// Mitsubishi GX Works2 project: v2(working)   PLC: FX3U/FX3UC

PROGRAM MAIN
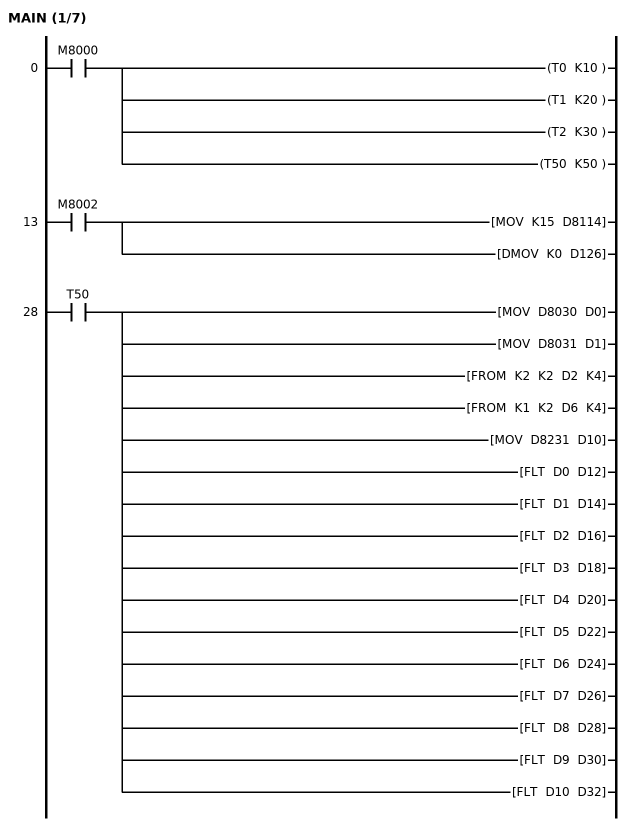
0     LD      M8000
      OUT     T0 K10
      OUT     T1 K20
      OUT     T2 K30
      OUT     T50 K50
13    LD      M8002
      MOV     K15 D8114
      DMOV    K0 D126
28    LD      T50
      MOV     D8030 D0
      MOV     D8031 D1
      FROM    K2 K2 D2 K4
      FROM    K1 K2 D6 K4
      MOV     D8231 D10
      FLT     D0 D12
      FLT     D1 D14
      FLT     D2 D16
      FLT     D3 D18
      FLT     D4 D20
      FLT     D5 D22
      FLT     D6 D24
      FLT     D7 D26
      FLT     D8 D28
      FLT     D9 D30
      FLT     D10 D32
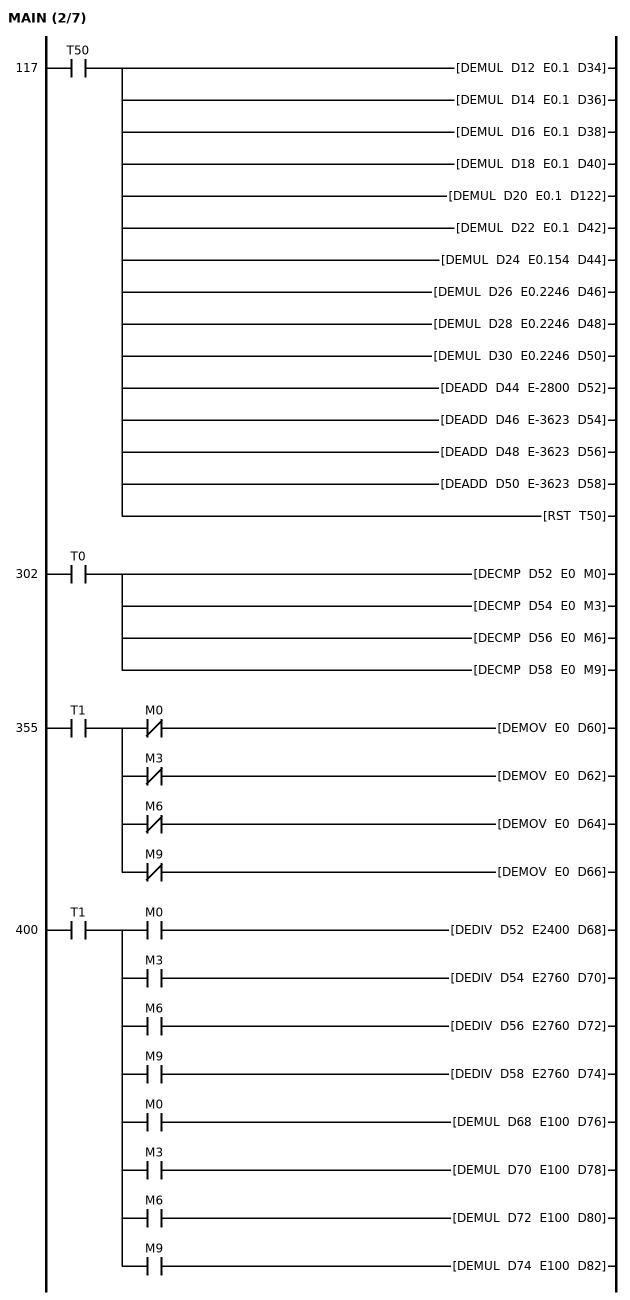
117   LD      T50
      DEMUL   D12 E0.1 D34
      DEMUL   D14 E0.1 D36
      DEMUL   D16 E0.1 D38
      DEMUL   D18 E0.1 D40
      DEMUL   D20 E0.1 D122
      DEMUL   D22 E0.1 D42
      DEMUL   D24 E0.154 D44
      DEMUL   D26 E0.2246 D46
      DEMUL   D28 E0.2246 D48
      DEMUL   D30 E0.2246 D50
      DEADD   D44 E-2800 D52
      DEADD   D46 E-3623 D54
      DEADD   D48 E-3623 D56
      DEADD   D50 E-3623 D58
      RST     T50
302   LD      T0
      DECMP   D52 E0 M0
      DECMP   D54 E0 M3
      DECMP   D56 E0 M6
      DECMP   D58 E0 M9
355   LD      T1
      MPS
      ANI     M0
      DEMOV   E0 D60
      MRD
      ANI     M3
      DEMOV   E0 D62
      MRD
      ANI     M6
      DEMOV   E0 D64
      MPP
      ANI     M9
      DEMOV   E0 D66
400   LD      T1
      MPS
      AND     M0
      DEDIV   D52 E2400 D68
      MRD
      AND     M3
      DEDIV   D54 E2760 D70
      MRD
      AND     M6
      DEDIV   D56 E2760 D72
      MRD
      AND     M9
      DEDIV   D58 E2760 D74
      MRD
      AND     M0
      DEMUL   D68 E100 D76
      MRD
      AND     M3
      DEMUL   D70 E100 D78
      MRD
      AND     M6
      DEMUL   D72 E100 D80
      MPP
      AND     M9
      DEMUL   D74 E100 D82
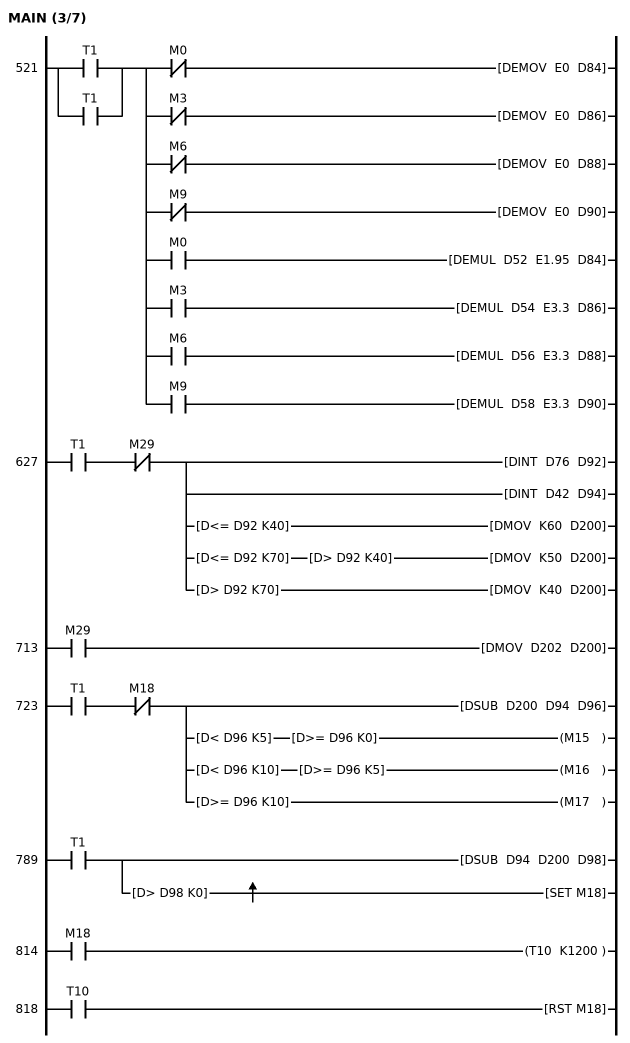
521   LD      T1
      OR      T1
      MPS
      ANI     M0
      DEMOV   E0 D84
      MRD
      ANI     M3
      DEMOV   E0 D86
      MRD
      ANI     M6
      DEMOV   E0 D88
      MRD
      ANI     M9
      DEMOV   E0 D90
      MRD
      AND     M0
      DEMUL   D52 E1.95 D84
      MRD
      AND     M3
      DEMUL   D54 E3.3 D86
      MRD
      AND     M6
      DEMUL   D56 E3.3 D88
      MPP
      AND     M9
      DEMUL   D58 E3.3 D90
627   LD      T1
      ANI     M29
      DINT    D76 D92
      DINT    D42 D94
      MPS
      ANDD<=  D92 K40
      DMOV    K60 D200
      MRD
      ANDD<=  D92 K70
      ANDD>   D92 K40
      DMOV    K50 D200
      MPP
      ANDD>   D92 K70
      DMOV    K40 D200
713   LD      M29
      DMOV    D202 D200
723   LD      T1
      ANI     M18
      DSUB    D200 D94 D96
      MPS
      ANDD<   D96 K5
      ANDD>=  D96 K0
      OUT     M15
      MRD
      ANDD<   D96 K10
      ANDD>=  D96 K5
      OUT     M16
      MPP
      ANDD>=  D96 K10
      OUT     M17
789   LD      T1
      DSUB    D94 D200 D98
      ANDD>   D98 K0
      MEP
      SET     M18
814   LD      M18
      OUT     T10 K1200
818   LD      T10
      RST     M18
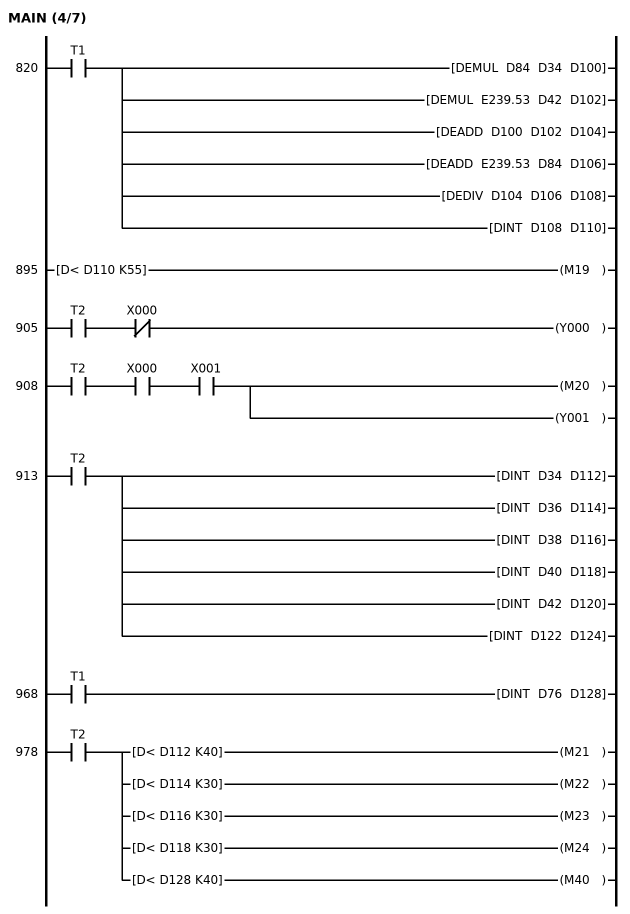
820   LD      T1
      DEMUL   D84 D34 D100
      DEMUL   E239.53 D42 D102
      DEADD   D100 D102 D104
      DEADD   E239.53 D84 D106
      DEDIV   D104 D106 D108
      DINT    D108 D110
895   LDD<    D110 K55
      OUT     M19
905   LD      T2
      ANI     X000
      OUT     Y000
908   LD      T2
      AND     X000
      AND     X001
      OUT     M20
      OUT     Y001
913   LD      T2
      DINT    D34 D112
      DINT    D36 D114
      DINT    D38 D116
      DINT    D40 D118
      DINT    D42 D120
      DINT    D122 D124
968   LD      T1
      DINT    D76 D128
978   LD      T2
      MPS
      ANDD<   D112 K40
      OUT     M21
      MRD
      ANDD<   D114 K30
      OUT     M22
      MRD
      ANDD<   D116 K30
      OUT     M23
      MRD
      ANDD<   D118 K30
      OUT     M24
      MPP
      ANDD<   D128 K40
      OUT     M40
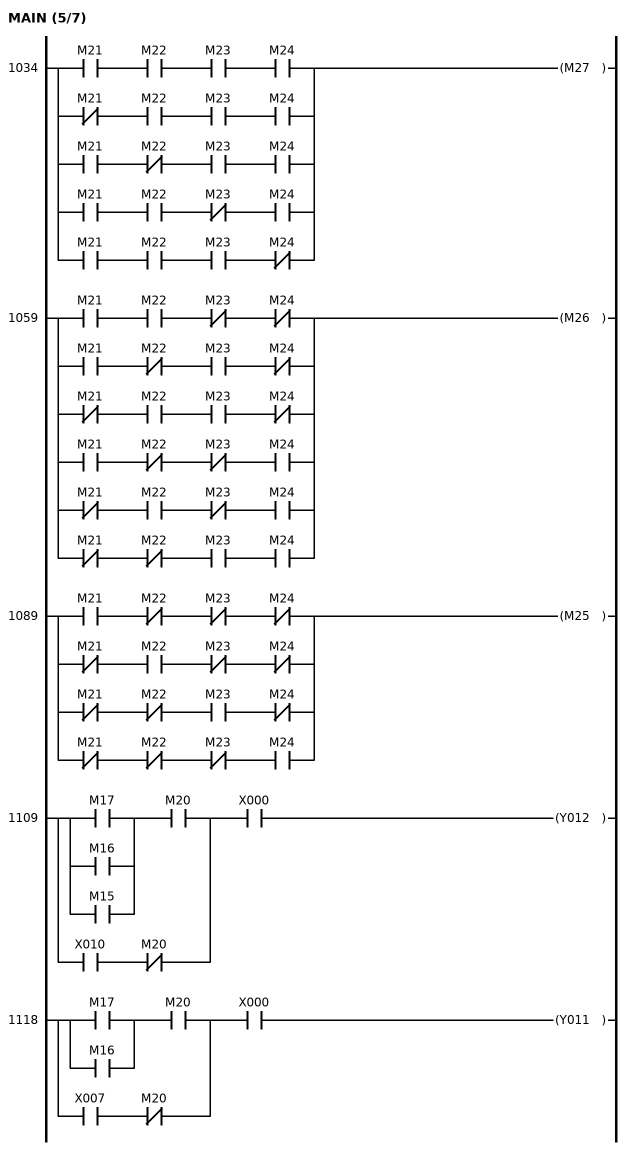
1034  LD      M21
      AND     M22
      AND     M23
      AND     M24
      LDI     M21
      AND     M22
      AND     M23
      AND     M24
      ORB
      LD      M21
      ANI     M22
      AND     M23
      AND     M24
      ORB
      LD      M21
      AND     M22
      ANI     M23
      AND     M24
      ORB
      LD      M21
      AND     M22
      AND     M23
      ANI     M24
      ORB
      OUT     M27
1059  LD      M21
      AND     M22
      ANI     M23
      ANI     M24
      LD      M21
      ANI     M22
      AND     M23
      ANI     M24
      ORB
      LDI     M21
      AND     M22
      AND     M23
      ANI     M24
      ORB
      LD      M21
      ANI     M22
      ANI     M23
      AND     M24
      ORB
      LDI     M21
      AND     M22
      ANI     M23
      AND     M24
      ORB
      LDI     M21
      ANI     M22
      AND     M23
      AND     M24
      ORB
      OUT     M26
1089  LD      M21
      ANI     M22
      ANI     M23
      ANI     M24
      LDI     M21
      AND     M22
      ANI     M23
      ANI     M24
      ORB
      LDI     M21
      ANI     M22
      AND     M23
      ANI     M24
      ORB
      LDI     M21
      ANI     M22
      ANI     M23
      AND     M24
      ORB
      OUT     M25
1109  LD      M17
      OR      M16
      OR      M15
      AND     M20
      LD      X010
      ANI     M20
      ORB
      AND     X000
      OUT     Y012
1118  LD      M17
      OR      M16
      AND     M20
      LD      X007
      ANI     M20
      ORB
      AND     X000
      OUT     Y011
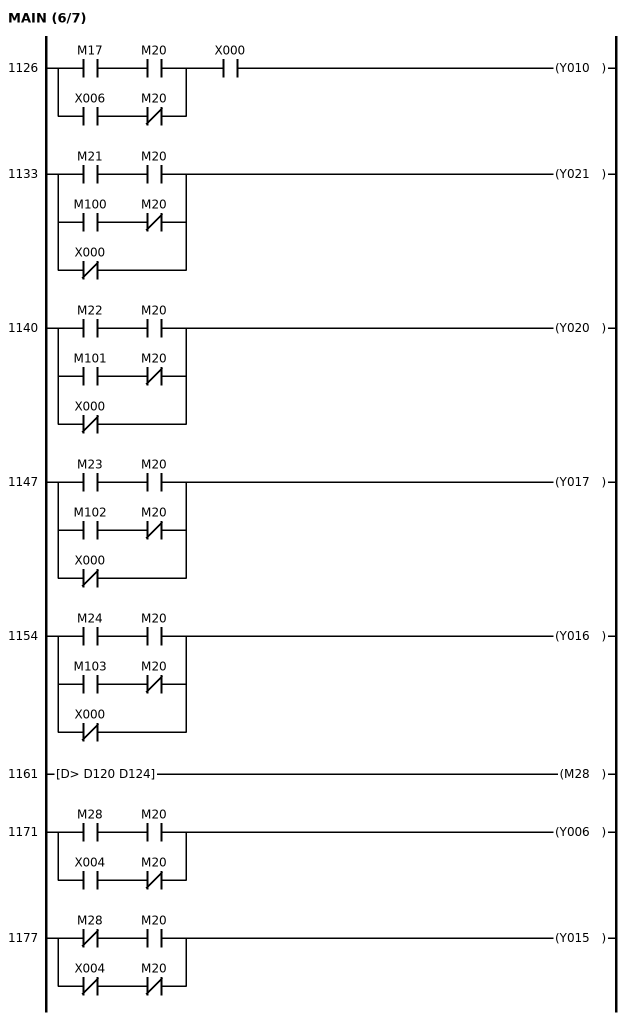
1126  LD      M17
      AND     M20
      LD      X006
      ANI     M20
      ORB
      AND     X000
      OUT     Y010
1133  LD      M21
      AND     M20
      LD      M100
      ANI     M20
      ORB
      ORI     X000
      OUT     Y021
1140  LD      M22
      AND     M20
      LD      M101
      ANI     M20
      ORB
      ORI     X000
      OUT     Y020
1147  LD      M23
      AND     M20
      LD      M102
      ANI     M20
      ORB
      ORI     X000
      OUT     Y017
1154  LD      M24
      AND     M20
      LD      M103
      ANI     M20
      ORB
      ORI     X000
      OUT     Y016
1161  LDD>    D120 D124
      OUT     M28
1171  LD      M28
      AND     M20
      LD      X004
      ANI     M20
      ORB
      OUT     Y006
1177  LDI     M28
      AND     M20
      LDI     X004
      ANI     M20
      ORB
      OUT     Y015
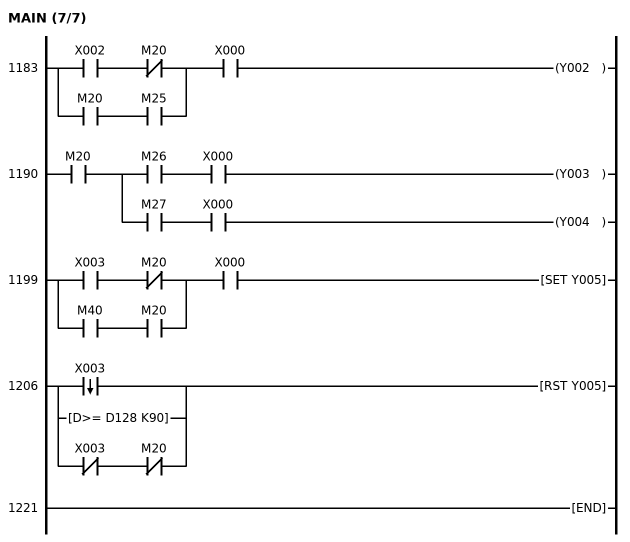
1183  LD      X002
      ANI     M20
      LD      M20
      AND     M25
      ORB
      AND     X000
      OUT     Y002
1190  LD      M20
      MPS
      AND     M26
      AND     X000
      OUT     Y003
      MPP
      AND     M27
      AND     X000
      OUT     Y004
1199  LD      X003
      ANI     M20
      LD      M40
      AND     M20
      ORB
      AND     X000
      SET     Y005
1206  LDF     X003
      ORD>=   D128 K90
      LDI     X003
      ANI     M20
      ORB
      RST     Y005
1221  END
END_PROGRAM
